(* IEC 61131-3 sources: kns-port-domestic/upstream/kns-pump-station/src/POUs/Model/FB_InflowProfile, 2 files *)

(* ---- FB_InflowProfile.decl.st ---- *)
// Назначение: суточный профиль притока: множитель f(tod) — линейная интерполяция точек профиля
//             (точка i — начало часа i, после 23 ч — снова точка 0), приток = rAverage_m3h · f.
//             Время суток приводится к [0, 24) по модулю; неконечное — как 0 ч. Среднее профиля
//             по умолчанию — 1,0: среднесуточный приток равен rAverage_m3h.
// Автор:      kr0nsch
// Версия:     0.1.0
// Документ:   docs/DESIGN.md, разделы 11.2, 11.3
FUNCTION_BLOCK FB_InflowProfile
VAR_INPUT
    rTimeOfDay_h : REAL;            // время суток модели, ч
    rAverage_m3h : REAL;            // средний приток (stSimCfg.rInflowAvg_m3h)
END_VAR
VAR_IN_OUT CONSTANT
    arProfile : ARRAY[0..GVL_Const.SIM_PROFILE_POINTS - 1] OF REAL;   // множители по часам (stSimCfg.arDailyProfile)
END_VAR
VAR_OUTPUT
    rFactor     : REAL;             // множитель профиля
    rInflow_m3h : REAL;             // приток по профилю, не меньше 0
END_VAR
VAR
    rTod_h   : REAL;                // время суток в [0, 24)
    rPos     : REAL;                // позиция в точках профиля
    diIndex  : DINT;                // точка слева
    uiLeft   : UINT;
    uiRight  : UINT;                // точка справа (по кругу)
END_VAR

(* ---- FB_InflowProfile.impl.st ---- *)
// 1. Время суток по модулю 24 ч (в том числе отрицательное)
IF PL.F_IsFinite(rIn := rTimeOfDay_h) THEN
    rTod_h := rTimeOfDay_h
              - GVL_Const.SIM_HOURS_PER_DAY * DINT_TO_REAL(TRUNC(rTimeOfDay_h / GVL_Const.SIM_HOURS_PER_DAY));
    IF rTod_h < 0.0 THEN
        rTod_h := rTod_h + GVL_Const.SIM_HOURS_PER_DAY;
    END_IF
    IF rTod_h >= GVL_Const.SIM_HOURS_PER_DAY THEN
        rTod_h := 0.0;
    END_IF
ELSE
    rTod_h := 0.0;
END_IF

// 2. Интерполяция между соседними точками; после последней — первая
rPos := rTod_h * UINT_TO_REAL(GVL_Const.SIM_PROFILE_POINTS) / GVL_Const.SIM_HOURS_PER_DAY;
diIndex := LIMIT(0, TRUNC(rPos), UINT_TO_DINT(GVL_Const.SIM_PROFILE_POINTS) - 1);
uiLeft := DINT_TO_UINT(diIndex);
uiRight := (uiLeft + 1) MOD GVL_Const.SIM_PROFILE_POINTS;
rFactor := arProfile[uiLeft] + (arProfile[uiRight] - arProfile[uiLeft]) * (rPos - DINT_TO_REAL(diIndex));

IF PL.F_IsFinite(rIn := rFactor) AND PL.F_IsFinite(rIn := rAverage_m3h) THEN
    rInflow_m3h := MAX(0.0, rAverage_m3h * rFactor);
ELSE
    rInflow_m3h := 0.0;
END_IF
